FUNCTION_BLOCK FB_Error
VAR_INPUT
	(* Input variables / Eingang Variablen *)
	bEnable					:BOOL;						(* Enable FB signal *)
	bReset					:BOOL;						(* Reset *)
	stAlarmIn					:ST_AlarmProperties;			(* Alarm output *)
END_VAR
VAR_OUTPUT
	(* Output variables / Ausgang Variablen *)
	stAlarmOut				:ST_AlarmProperties;			(* Alarm output *)
END_VAR
VAR_IN_OUT

END_VAR
VAR
	(* Enummerations *)

	(* Variables *)

	(* References *)

	(* Interfaces *)

	(* Instances *)

END_VAR

(* Check method enabled *)
IF NOT bEnable
THEN
	RETURN;
END_IF;

IF bReset
THEN
	IF stAlarmOut.bActive
	THEN
		stAlarmOut.bActive := FALSE;
		(*stAlarmOut.enType := ET_AlarmType_eIdle;*)
		(*stAlarmOut.dtDateTime := DT#1970-01-01-00:00;*)
		(*stAlarmOut.dnCode := 0;*)
	END_IF;
ELSE
	IF stAlarmIn.bActive
	    AND NOT stAlarmOut.bActive
	THEN
		stAlarmOut.bActive := TRUE;
		stAlarmOut.enType := stAlarmIn.enType;
		stAlarmOut.dtDateTime := stAlarmIn.dtDateTime;
		stAlarmOut.dnCode := stAlarmIn.dnCode;
	END_IF;
END_IF;

END_FUNCTION_BLOCK

(* stored: Version 1.1.0.1, ProductVersion 3.1.4024.15
   POU FB_Error: Id {ce39f4f3-c641-47db-b1ea-613c4068ce62}, SpecialFunc None *)
